Omron CX-Programmer project OmronTeachingExample (CX-Programmer 9.75)

# PLC ExamplePLC: CP1L L

## Program Main (cyclic task 0)

### Section Section1

### Section Instruction_Probe

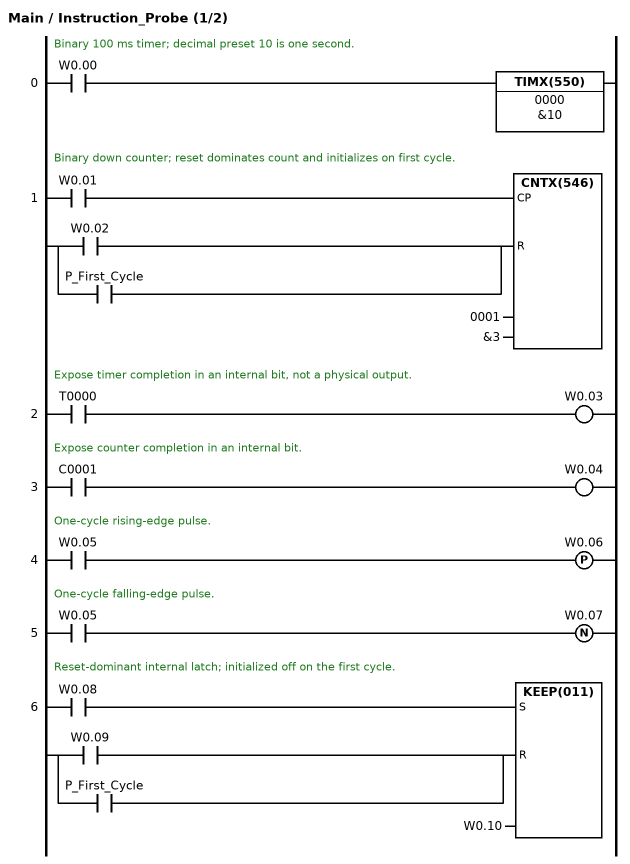
; rung 0: Binary 100 ms timer; decimal preset 10 is one second.
LD W0.00
TIMX(550) 0000 &10
; rung 1: Binary down counter; reset dominates count and initializes on first cycle.
LD W0.01
LD W0.02
OR P_First_Cycle
CNTX(546) 0001 &3
; rung 2: Expose timer completion in an internal bit, not a physical output.
LD T0000
OUT W0.03
; rung 3: Expose counter completion in an internal bit.
LD C0001
OUT W0.04
; rung 4: One-cycle rising-edge pulse.
LD W0.05
DIFU(013) W0.06
; rung 5: One-cycle falling-edge pulse.
LD W0.05
DIFD(014) W0.07
; rung 6: Reset-dominant internal latch; initialized off on the first cycle.
LD W0.08
LD W0.09
OR P_First_Cycle
KEEP(011) W0.10

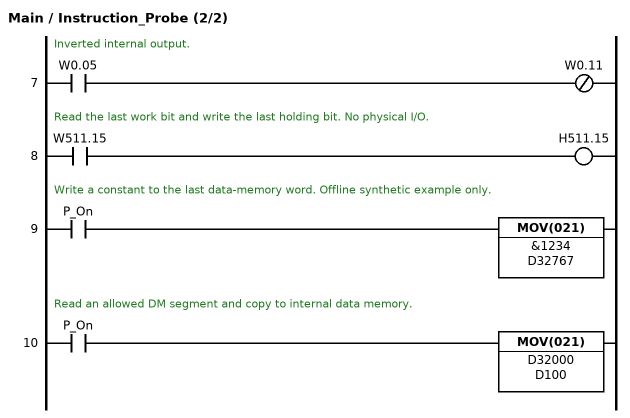
; rung 7: Inverted internal output.
LD W0.05
OUTNOT W0.11
; rung 8: Read the last work bit and write the last holding bit. No physical I/O.
LD W511.15
OUT H511.15
; rung 9: Write a constant to the last data-memory word. Offline synthetic example only.
LD P_On
MOV(021) &1234 D32767
; rung 10: Read an allowed DM segment and copy to internal data memory.
LD P_On
MOV(021) D32000 D100

### Section END
; rung 0
END(001)